    rq_activate_all_grippers(True)
    # end: URCap Program Node
  end
  $ 57 "zero_ftsensor()"
  zero_ftsensor()
  $ 58 "EXTT"
  $ 59 "Set GRP_3F_Enable=Off"
  set_standard_digital_out(4, False)
  $ 60 "Set DO[6]=Off"
  set_standard_digital_out(6, False)
  $ 61 "Set GRP_3F_Decap=Off"
  set_standard_digital_out(3, False)
  $ 62 "Set GRP_3F_Cap=Off"
  set_standard_digital_out(2, False)
  $ 63 "Set GRP_3F_Open=Off"
  set_standard_digital_out(5, False)
  $ 64 "PSE_T≔get_tool_free_pose(dir=[0,0,0.150], move_in_base_frame=True)"
  global PSE_T=get_tool_free_pose(dir=[0,0,0.150], move_in_base_frame=True)
  $ 65 "If is_reachable(Base_const, [PSE_T])"
  if (is_reachable(p[0.0,0.0,0.0,0.0,0.0,0.0], [PSE_T])):
    $ 66 "MoveL"
    $ 67 "PSE_T" "breakAfter"
    movel(PSE_T, a=1.2, v=0.15)
  end
  $ 68 "powder dispensing variable init"
  $ 69 "Start_thread≔ False "
  global Start_thread=  False
  $ 70 "vib_mot_thread≔ False "
  global vib_mot_thread=  False
  $ 71 "kp≔0.0002"
  global kp=0.0002
  $ 72 "ki≔0.001"
  global ki=0.001
  $ 73 "kd≔0.01"
  global kd=0.01
  $ 74 "dt≔0.05"
  global dt=0.05
  $ 75 "Integral_error≔0"
  global Integral_error=0
  $ 76 "current_error≔0"
  global current_error=0
  $ 77 "previous_error≔0"
  global previous_error=0
  $ 78 "tilt_increment≔0"
  global tilt_increment=0
  $ 79 "tilt_angle≔-1"
  global tilt_angle=-1
  $ 80 "diff≔0"
  global diff=0
  $ 81 "current_pose≔get_actual_tcp_pose()"
  global current_pose= get_actual_tcp_pose ()
  $ 896 "Thread_1"
  thread Thread_1():
    while (True):
      $ 897 "If Start_thread≟ True "
      if (Start_thread ==   True  ):
        $ 898 "Weight_value≔get_weight()"
        global Weight_value=get_weight()
        $ 899 "sync()"
        sync()
      end
    end
  end
  threadId_Thread_1 = run Thread_1()
  $ 900 "Thread_2"
  thread Thread_2():
    while (True):
      $ 901 "Loop vib_mot_thread≟ True "
      thread Thread_while_901():
        while (True):
          $ 902 "diff≔Target_weight-Weight_value"
          global diff=Target_weight-Weight_value
          $ 903 "If diff>0.08"
          global thread_flag_903=0
          thread Thread_if_903():
            $ 904 "Set AO[0]=4.0"
            set_standard_analog_out(0, 0.4)
            thread_flag_903 = 1
          end
          if (diff>0.08):
            global thread_handler_903=run Thread_if_903()
            while (thread_flag_903 == 0):
              if not(diff>0.08):
                kill thread_handler_903
                thread_flag_903 = 2
              else:
                sync()
              end
            end
          else:
            thread_flag_903 = 2
          end
          if (thread_flag_903 == 2):
            $ 905 "ElseIf diff≥0.04 and diff≤0.08"
            global thread_flag_905=0
            thread Thread_if_905():
              $ 906 "vibration_1()"
              vibration_1()
              thread_flag_905 = 1
            end
            if (diff >= 0.04 and diff <= 0.08):
              global thread_handler_905=run Thread_if_905()
              while (thread_flag_905 == 0):
                if not(diff >= 0.04 and diff <= 0.08):
                  kill thread_handler_905
                  thread_flag_905 = 2
                else:
                  sync()
                end
              end
            else:
              thread_flag_905 = 2
            end
            if (thread_flag_905 == 2):
              $ 907 "ElseIf diff≥0.01 and diff<0.04"
              if (diff >= 0.01 and diff<0.04):
                $ 908 "vibration_2()"
                vibration_2()
              else:
                $ 909 "ElseIf diff>0 and diff<0.01"
                if (diff>0 and diff<0.01):
                  $ 910 "vibration_3()"
                  vibration_3()
                else:
                  $ 911 "Else" "noBreak"
                  $ 912 "Set AO[0]=0.0"
                  set_standard_analog_out(0, 0.0)
                end
              end
            end
          end
        end
      end
      if (vib_mot_thread ==   True  ):
        global thread_handler_901=run Thread_while_901()
        while (vib_mot_thread ==   True  ):
          sync()
        end
        kill thread_handler_901
      end
      $ 915 "sync()"
      sync()
    end
  end
  threadId_Thread_2 = run Thread_2()
  while (True):
    $ 82 "Robot Program"
    $ 83 "MAIN"
    $ 84 "command_manager(external_control='uGO', cond_suspend=(ITM_Manipulated and AMR_AtTarget and AMR_Charging and AMR_Battery<40), cond_unsuspend=(AMR_Battery≟60))"
    command_manager(external_control="uGO", cond_suspend=(ITM_Manipulated  and  AMR_AtTarget  and  AMR_Charging  and  AMR_Battery<40), cond_unsuspend=(AMR_Battery == 60))
    $ 85 "log_state(STATE_Info)"
    log_state(STATE_Info)
    $ 86 "Switch STATE"
    switch_1 = STATE
    $ 87 "Case 1"
    if (1 == switch_1):
      $ 88 "Stopping"
      $ 89 "STATE_Info≔'Stopping'"
      global STATE_Info="Stopping"
      $ 90 "end_freedrive_mode()"
      end_freedrive_mode()
      $ 91 "Set"
      set_tcp(p[0.0,0.0,0.161,3.1415,0.0,0.0])
      $ 92 "PSE_T≔get_tool_free_pose(dir=[0,0,0.150], move_in_base_frame=True)"
      global PSE_T=get_tool_free_pose(dir=[0,0,0.150], move_in_base_frame=True)
      $ 93 "If is_reachable(Base_const, [PSE_T])"
      if (is_reachable(p[0.0,0.0,0.0,0.0,0.0,0.0], [PSE_T])):
        $ 94 "MoveL"
        $ 95 "PSE_T" "breakAfter"
        movel(PSE_T, a=1.2, v=0.15)
      end
      $ 96 "do_transition(keep_rxry=OBJ_Picked, r=0)"
      do_transition(keep_rxry=OBJ_Picked, r=0)
      $ 105 "Call Sub_AMR_MiR_V3"
      Sub_AMR_MiR_V3()
      $ 106 "If stopping() and AMR_Done"
      if (stopping()  and  AMR_Done):
        $ 107 "STATE≔2"
        global STATE=2
        $ 108 "ugo_update_outputs()"
        ugo_update_outputs()
      end
    elif (2 == switch_1):
      $ 109 "Case 2"
      $ 110 "Stopped"
      $ 111 "STATE_Info≔'Stopped'"
      global STATE_Info="Stopped"
      $ 112 "Call Sub_AMR_MiR_V3"
      Sub_AMR_MiR_V3()
      $ 113 "If CMD_Reset"
      if (CMD_Reset):
        $ 114 "STATE≔3"
        global STATE=3
        $ 115 "ugo_update_outputs()"
        ugo_update_outputs()
      end
    elif (3 == switch_1):
      $ 116 "Case 3"
      $ 117 " Resetting"
      $ 118 "STATE_Info≔'Resetting'"
      global STATE_Info="Resetting"
      $ 119 "uML"
      $ 120 "reset_error()"
      reset_error()
      $ 121 "reset_warning()"
      reset_warning()
      $ 122 "PROCESS_Step≔0"
      global PROCESS_Step=0
      $ 123 "PROCESS_Info≔''"
      global PROCESS_Info=""
      $ 124 "ARM_Referenced≔ False "
      global ARM_Referenced=  False
      $ 125 "WRK_Done≔ False "
      global WRK_Done=  False
      $ 126 "ITM_Prepared≔ False "
      global ITM_Prepared=  False
      $ 127 "ITM_Manipulated≔ False "
      global ITM_Manipulated=  False
      $ 128 "STP≔0"
      global STP=0
      $ 129 "Action≔0"
      global Action=0
      $ 130 "Action_Info≔''"
      global Action_Info=""
      $ 131 "ITM_ID≔0"
      global ITM_ID=0
      $ 132 "JIG≔0"
      global JIG=0
      $ 133 "JIG_Slot≔0"
      global JIG_Slot=0
      $ 134 "Task_info≔''"
      global Task_info=""
      $ 135 "Set"
      set_tcp(p[0.0,0.0,0.161,3.1415,0.0,0.0])
      $ 136 "App"
      $ 137 "'ADD APPLICATION SPECIFIC COMMANDS'"
      # 'ADD APPLICATION SPECIFIC COMMANDS'
      $ 138 "OBJ_Type≔0"
      global OBJ_Type=0
      $ 139 "OBJ_Nbr≔0"
      global OBJ_Nbr=0
      $ 140 "If CNT_Rack_Output≥50"
      if (CNT_Rack_Output >= 50):
        $ 141 "CNT_Rack_Output≔0"
        global CNT_Rack_Output=0
      end
      $ 142 "TASK≔struct(ID=0, NAVI=struct(target=0, footprint=0, protectiveOff=0, dock=0), WORK=struct(ITM_ID_Src=0, JIG_ID_Src=0, OBJ_Nbr_Src=0, ACT_Src=0, ITM_ID_Tgt=0, JIG_ID_Tgt=0, OBJ_Nbr_Tgt=0, ACT_Tgt=0, OBJ_Type=0))"
      global TASK=struct(ID=0, NAVI=struct(target=0, footprint=0, protectiveOff=0, dock=0), WORK=struct(ITM_ID_Src=0, JIG_ID_Src=0, OBJ_Nbr_Src=0, ACT_Src=0, ITM_ID_Tgt=0, JIG_ID_Tgt=0, OBJ_Nbr_Tgt=0, ACT_Tgt=0, OBJ_Type=0))
      $ 143 "Call Sub_AMR_MiR_V3"
      Sub_AMR_MiR_V3()
      $ 144 "If resetting() and AMR_Done"
      if (resetting()  and  AMR_Done):
        $ 145 "STATE≔4"
        global STATE=4
        $ 146 "ugo_update_outputs()"
        ugo_update_outputs()
      end
    elif (4 == switch_1):
      $ 147 "Case 4"
      $ 148 "Idle"
      $ 149 "STATE_Info≔'Idle'"
      global STATE_Info="Idle"
      $ 150 "If CMD_Start"
      if (CMD_Start):
        $ 151 "STATE≔5"
        global STATE=5
        $ 152 "ugo_update_outputs()"
        ugo_update_outputs()
      end
    elif (5 == switch_1):
      $ 153 "Case 5"
      $ 154 "Starting"
      $ 155 "STATE_Info≔'Starting'"
      global STATE_Info="Starting"
      $ 156 "'ADD COMMANDS WHAT TO START WITH'"
      # 'ADD COMMANDS WHAT TO START WITH'
      $ 157 "Call Sub_AMR_MiR_V3"
      Sub_AMR_MiR_V3()
      $ 158 "get ugo data"
      $ 159 "Assign Tasks"
      $ 160 "TASK.ID = ugo_get_task()"
      TASK.ID = ugo_get_task()
      $ 161 "If TASK.ID≟1"
      if (TASK.ID == 1):
        $ 162 "Task_info≔'Charge'"
        global Task_info="Charge"
        $ 163 "Parameters"
        $ 164 "AMR_PosTarget≔1"
        global AMR_PosTarget=1
      else:
        $ 165 "ElseIf TASK.ID≟9"
        if (TASK.ID == 9):
          $ 166 "'Pick Sarstedt Rack from Variable source'"
          # 'Pick Sarstedt Rack from Variable source'
          $ 167 "Task_info≔'Navigate to Target'"
          global Task_info="Navigate to Target"
          $ 168 "Parameters"
          $ 169 "AMR_PosTarget≔UGO.read_input('00','ITM_ID')"
          global AMR_PosTarget=UGO.read_input("00","ITM_ID")
        else:
          $ 170 "ElseIf TASK.ID≟10"
          if (TASK.ID == 10):
            $ 171 "'Pick Sarstedt Rack from Variable source'"
            # 'Pick Sarstedt Rack from Variable source'
            $ 172 "Task_info≔'Pick Rack'"
            global Task_info="Pick Rack"
            $ 173 "AMR_PosTarget≔2"
            global AMR_PosTarget=2
            $ 174 "Parameters"
            $ 175 "ITM_ID≔UGO.read_input('00','ITM_ID')"
            global ITM_ID=UGO.read_input("00","ITM_ID")
            $ 176 "JIG≔UGO.read_input('00','JIG_ID')"
            global JIG=UGO.read_input("00","JIG_ID")
            $ 177 "OBJ_Type≔3"
            global OBJ_Type=3
          else:
            $ 178 "ElseIf TASK.ID≟11"
            if (TASK.ID == 11):
              $ 179 "'Place Sarstedt Rack on Variable target'"
              # 'Place Sarstedt Rack on Variable target'
              $ 180 "Task_info≔'Place Rack'"
              global Task_info="Place Rack"
              $ 181 "AMR_PosTarget≔2"
              global AMR_PosTarget=2
              $ 182 "Parameters"
              $ 183 "ITM_ID≔UGO.read_input('00','ITM_ID')"
              global ITM_ID=UGO.read_input("00","ITM_ID")
              $ 184 "JIG≔UGO.read_input('00','JIG_ID')"
              global JIG=UGO.read_input("00","JIG_ID")
              $ 185 "OBJ_Type≔3"
              global OBJ_Type=3
            else:
              $ 187 "ElseIf TASK.ID≟12"
              if (TASK.ID == 12):
                $ 188 "Task_info≔'Decapping'"
                global Task_info="Decapping"
                $ 189 "Parameters"
                $ 190 "ITM_ID≔1"
                global ITM_ID=1
                $ 191 "AMR_PosTarget≔AMR_PosActual"
                global AMR_PosTarget=AMR_PosActual
                $ 192 "PRC_TubCounter≔0"
                global PRC_TubCounter=0
              else:
                $ 193 "ElseIf TASK.ID≟13"
                if (TASK.ID == 13):
                  $ 194 "Task_info≔'Empty racks'"
                  global Task_info="Empty racks"
                  $ 195 "Parameters"
                  $ 196 "ITM_ID≔1"
                  global ITM_ID=1
                  $ 197 "AMR_PosTarget≔AMR_PosActual"
                  global AMR_PosTarget=AMR_PosActual
                else:
                  $ 198 "ElseIf TASK.ID≟16"
                  if (TASK.ID == 16):
                    $ 199 "Task_info≔'Decap + Barcode'"
                    global Task_info="Decap + Barcode"
                    $ 200 "Parameters"
                    $ 202 "OBJs_String≔UGO.read_input('00','ObjPos')"
                    global OBJs_String=UGO.read_input("00","ObjPos")
                    $ 203 "OBJs_List≔make_list(length = elements_in_string(OBJs_String), initial_value = -1, capacity = 50)"
                    global OBJs_List=make_list(length = elements_in_string(OBJs_String), initial_value = -1, capacity = 50)
                    $ 204 "OBJs_List≔string_to_list(OBJs_String)"
                    global OBJs_List=string_to_list(OBJs_String)
                    $ 205 "ITM_ID≔1"
                    global ITM_ID=1
                    $ 206 "OBJ_Type≔2"
                    global OBJ_Type=2
                    $ 207 "JIG≔7"
                    global JIG=7
                    $ 208 "AMR_PosTarget≔AMR_PosActual"
                    global AMR_PosTarget=AMR_PosActual
                  else:
                    $ 209 "ElseIf TASK.ID≟30"
                    if (TASK.ID == 30):
                      $ 210 "Task_info≔'Getting bottles'"
                      global Task_info="Getting bottles"
                      $ 211 "Parameters"
                      $ 212 "ITM_ID≔1"
                      global ITM_ID=1
                      $ 213 "OBJ_Type≔4"
                      global OBJ_Type=4
                      $ 214 "JIG≔9"
                      global JIG=9
                      $ 215 "AMR_PosTarget≔4"
                      global AMR_PosTarget=4
                    else:
                      $ 216 "ElseIf TASK.ID≟40"
                      if (TASK.ID == 40):
                        $ 217 "Task_info≔'Placing bottles'"
                        global Task_info="Placing bottles"
                        $ 218 "Parameters"
                        $ 219 "ITM_ID≔1"
                        global ITM_ID=1
                        $ 220 "OBJ_Type≔4"
                        global OBJ_Type=4
                        $ 221 "JIG≔10"
                        global JIG=10
                        $ 222 "AMR_PosTarget≔4"
                        global AMR_PosTarget=4
                      else:
                        $ 223 "ElseIf TASK.ID≟41"
                        if (TASK.ID == 41):
                          $ 224 "Task_info≔'Shaking bottle'"
                          global Task_info="Shaking bottle"
                          $ 225 "Parameters"
                          $ 226 "ITM_ID≔1"
                          global ITM_ID=1
                          $ 227 "OBJ_Type≔4"
                          global OBJ_Type=4
                          $ 228 "JIG≔11"
                          global JIG=11
                          $ 229 "AMR_PosTarget≔4"
                          global AMR_PosTarget=4
                        else:
                          $ 230 "ElseIf TASK.ID≟42"
                          if (TASK.ID == 42):
                            $ 231 "Task_info≔'Decap the bottle'"
                            global Task_info="Decap the bottle"
                            $ 232 "Parameters"
                            $ 233 "ITM_ID≔1"
                            global ITM_ID=1
                            $ 234 "OBJ_Type≔4"
                            global OBJ_Type=4
                            $ 235 "AMR_PosTarget≔4"
                            global AMR_PosTarget=4
                          else:
                            $ 236 "ElseIf TASK.ID≟43"
                            if (TASK.ID == 43):
                              $ 237 "Task_info≔'Pick the Rack'"
                              global Task_info="Pick the Rack"
                              $ 238 "AMR_PosTarget≔5"
                              global AMR_PosTarget=5
                              $ 239 "Parameters"
                              $ 240 "ITM_ID≔UGO.read_input('00','ITM_ID')"
                              global ITM_ID=UGO.read_input("00","ITM_ID")
                              $ 241 "JIG≔UGO.read_input('00','JIG_ID')"
                              global JIG=UGO.read_input("00","JIG_ID")
                              $ 242 "OBJ_Type≔3"
                              global OBJ_Type=3
                            else:
                              $ 243 "ElseIf TASK.ID≟45"
                              if (TASK.ID == 45):
                                $ 244 "Task_info≔'pick the Vial'"
                                global Task_info="pick the Vial"
                                $ 245 "Parameters"
                                $ 246 "ITM_ID≔1"
                                global ITM_ID=1
                                $ 247 "OBJ_Type≔4"
                                global OBJ_Type=4
                                $ 248 "JIG≔12"
                                global JIG=12
                                $ 249 "AMR_PosTarget≔5"
                                global AMR_PosTarget=5
                              else:
                                $ 250 "ElseIf TASK.ID≟46"
                                if (TASK.ID == 46):
                                  $ 251 "Task_info≔'Decap the Vial'"
                                  global Task_info="Decap the Vial"
                                  $ 252 "Parameters"
                                  $ 253 "ITM_ID≔1"
                                  global ITM_ID=1
                                  $ 254 "OBJ_Type≔4"
                                  global OBJ_Type=4
                                  $ 255 "JIG≔13"
                                  global JIG=13
                                  $ 256 "AMR_PosTarget≔5"
                                  global AMR_PosTarget=5
                                else:
                                  $ 257 "ElseIf TASK.ID≟47"
                                  if (TASK.ID == 47):
                                    $ 258 "Task_info≔'Liquid Transfer'"
                                    global Task_info="Liquid Transfer"
                                    $ 259 "Parameters"
                                    $ 260 "ITM_ID≔1"
                                    global ITM_ID=1
                                    $ 261 "OBJ_Type≔4"
                                    global OBJ_Type=4
                                    $ 262 "JIG≔14"
                                    global JIG=14
                                    $ 263 "AMR_PosTarget≔3"
                                    global AMR_PosTarget=3
                                  else:
                                    $ 264 "ElseIf TASK.ID≟48"
                                    if (TASK.ID == 48):
                                      $ 265 "Task_info≔'Place_rack'"
                                      global Task_info="Place_rack"
                                      $ 266 "Parameters"
                                      $ 267 "ITM_ID≔1"
                                      global ITM_ID=1
                                      $ 268 "OBJ_Type≔3"
                                      global OBJ_Type=3
                                      $ 269 "JIG≔7"
                                      global JIG=7
                                      $ 270 "AMR_PosTarget≔5"
                                      global AMR_PosTarget=5
                                    else:
                                      $ 271 "ElseIf TASK.ID≟49"
                                      if (TASK.ID == 49):
                                        $ 272 "Task_info≔'Pick Containers'"
                                        global Task_info="Pick Containers"
                                        $ 273 "Parameters"
                                        $ 274 "ITM_ID≔1"
                                        global ITM_ID=1
                                        $ 275 "OBJ_Type≔6"
                                        global OBJ_Type=6
                                        $ 276 "JIG≔15"
                                        global JIG=15
                                        $ 277 "AMR_PosTarget≔3"
                                        global AMR_PosTarget=3
                                      else:
                                        $ 278 "ElseIf TASK.ID≟50"
                                        if (TASK.ID == 50):
                                          $ 279 "Task_info≔'Decap Containers'"
                                          global Task_info="Decap Containers"
                                          $ 280 "Parameters"
                                          $ 281 "ITM_ID≔1"
                                          global ITM_ID=1
                                          $ 282 "OBJ_Type≔6"
                                          global OBJ_Type=6
                                          $ 283 "JIG≔16"
                                          global JIG=16
                                          $ 284 "AMR_PosTarget≔5"
                                          global AMR_PosTarget=5
                                        else:
                                          $ 285 "ElseIf TASK.ID≟51"
                                          if (TASK.ID == 51):
                                            $ 286 "Task_info≔'Detect Spatula and transfer powder'"
                                            global Task_info="Detect Spatula and transfer powder"
                                            $ 287 "Parameters"
                                            $ 288 "ITM_ID≔1"
                                            global ITM_ID=1
                                            $ 289 "Target_weight≔(UGO.read_input('00','Target_weight'))/1000"
                                            global Target_weight=(UGO.read_input("00","Target_weight"))/1000
                                            $ 290 "OBJ_Type≔8"
                                            global OBJ_Type=8
                                            $ 291 "JIG≔16"
                                            global JIG=16
                                            $ 292 "AMR_PosTarget≔5"
                                            global AMR_PosTarget=5
                                          else:
                                            $ 293 "ElseIf TASK.ID≟99"
                                            if (TASK.ID == 99):
                                              $ 294 "Task_info≔'Decapping and barcode alignment'"
                                              global Task_info="Decapping and barcode alignment"
                                              $ 295 "Parameters"
                                              $ 296 "PRC_TubNumber≔UGO.read_input('00','TubesNb')"
                                              global PRC_TubNumber=UGO.read_input("00","TubesNb")
                                              $ 297 "PRC_TubCounter≔0"
                                              global PRC_TubCounter=0
                                              $ 298 "ITM_ID≔1"
                                              global ITM_ID=1
                                              $ 299 "AMR_PosTarget≔AMR_PosActual"
                                              global AMR_PosTarget=AMR_PosActual
                                            else:
                                              $ 334 "Else" "noBreak"
                                              $ 335 "set_error(ERROR_WRONG_ORDER)"
                                              set_error(ERROR_WRONG_ORDER)
                                            end
                                          end
                                        end
                                      end
                                    end
                                  end
                                end
                              end
                            end
                          end
                        end
                      end
                    end
                  end
                end
              end
            end
          end
        end
      end
      $ 336 "test ugo"
      $ 337 "Wait: 0.2"
      sleep(0.2)
      $ 338 "ugo_update_outputs()"
      ugo_update_outputs()
      $ 339 "If starting() and AMR_Done"
      if (starting()  and  AMR_Done):
        $ 340 "log_message(Task_info, 'New Task: ')"
        log_message(Task_info, "New Task: ")
        $ 341 "log_message(to_str(TASK.ID), 'Task_ID: ')"
        log_message(to_str(TASK.ID), "Task_ID: ")
        $ 342 "do_transition(keep_rxry=OBJ_Picked)"
        do_transition(keep_rxry=OBJ_Picked)
        $ 343 "STATE≔6"
        global STATE=6
        $ 344 "ugo_update_outputs()"
        ugo_update_outputs()
      end
    elif (6 == switch_1):
      $ 345 "Case 6"
      $ 346 "Execute"
      $ 347 "STATE_Info≔'Execute'"
      global STATE_Info="Execute"
      $ 348 "If  not CMD_Hold and not CMD_Suspend"
      global thread_flag_348=0
      thread Thread_if_348():
        $ 349 "Switch PROCESS_Step"
        switch_2 = PROCESS_Step
        $ 350 "Case 0"
        if (0 == switch_2):
          $ 351 "PROCESS_Info≔'process control'"
          global PROCESS_Info="process control"
          $ 352 "log_process(PROCESS_Info)"
          log_process(PROCESS_Info)
          $ 353 "process control"
          $ 354 "If  not AMR_AtTarget"
          if (  not  AMR_AtTarget):
            $ 355 "PROCESS_Step≔1"
            global PROCESS_Step=1
          else:
            $ 356 "ElseIf (( not ITM_Prepared and  not WRK_Done) or (ITM_Prepared and WRK_Done))"
            if (((  not  ITM_Prepared  and    not  WRK_Done)  or  (ITM_Prepared  and  WRK_Done))):
              $ 357 "PROCESS_Step≔2"
              global PROCESS_Step=2
            else:
              $ 358 "ElseIf  not WRK_Done"
              if (  not  WRK_Done):
                $ 359 "PROCESS_Step≔3"
                global PROCESS_Step=3
              else:
                $ 360 "Else" "noBreak"
                $ 361 "task finished"
                $ 362 "PROCESS_Info≔''"
                global PROCESS_Info=""
                $ 363 "STATE≔7"
                global STATE=7
                $ 364 "ugo_update_outputs()"
                ugo_update_outputs()
              end
            end
          end
        elif (1 == switch_2):
          $ 365 "Case 1"
          $ 366 "navigate"
          $ 367 "'MOVING THE uML'"
          # 'MOVING THE uML'
          $ 368 "PROCESS_Info≔'move to target'"
          global PROCESS_Info="move to target"
          $ 369 "log_process(PROCESS_Info)"
          log_process(PROCESS_Info)
          $ 370 "If TASK.ID≟1"
          if (TASK.ID == 1):
            $ 371 "Action≔51"
            global Action=51
          else:
            $ 372 "Else" "noBreak"
            $ 373 "Action≔52"
            global Action=52
          end
          $ 374 "Call Sub_AMR_MiR_V3"
          Sub_AMR_MiR_V3()
          $ 375 "If AMR_Done"
          if (AMR_Done):
            $ 376 "PROCESS_Step≔0"
            global PROCESS_Step=0
          end
        elif (2 == switch_2):
          $ 377 "Case 2"
          $ 378 "prepare"
          $ 379 "'THINGS THAT HAVE TO BE DONE ONCE IN A SEQUENCE,WORKFLOW'"
          # 'THINGS THAT HAVE TO BE DONE ONCE IN A SEQUENCE,WORKFLOW'
          $ 380 "PROCESS_Info≔'prepare for work'"
          global PROCESS_Info="prepare for work"
          $ 381 "log_process(PROCESS_Info)"
          log_process(PROCESS_Info)
          $ 382 "If TASK.WORK.ITM_ID_Src>1"
          if (TASK.WORK.ITM_ID_Src>1):
            $ 383 "ITM_ID≔TASK.WORK.ITM_ID_Src"
            global ITM_ID=TASK.WORK.ITM_ID_Src
          else:
            $ 384 "ElseIf TASK.WORK.ITM_ID_Tgt>1"
            if (TASK.WORK.ITM_ID_Tgt>1):
              $ 385 "ITM_ID≔TASK.WORK.ITM_ID_Tgt"
              global ITM_ID=TASK.WORK.ITM_ID_Tgt
            end
          end
          $ 386 "If  not ARM_Referenced and (ITM_ID≠0)"
          if (  not  ARM_Referenced  and  (ITM_ID != 0)):
            $ 387 "STP≔1"
            global STP=1
          else:
            $ 388 "ElseIf ARM_Referenced or (ITM_ID≟0)"
            if (ARM_Referenced  or  (ITM_ID == 0)):
              $ 389 "STP≔2"
              global STP=2
            end
          end
          $ 390 "Switch STP"
          switch_3 = STP
          $ 391 "Case 1"
          if (1 == switch_3):
            $ 392 "reference"
            $ 393 "STP_Info≔'reference at target position'"
            global STP_Info="reference at target position"
            $ 394 "log_step(STP_Info)"
            log_step(STP_Info)
            $ 395 "If ITM_ID≟1"
            if (ITM_ID == 1):
              $ 396 "CAM_Done≔ True "
              global CAM_Done=  True
            else:
              $ 397 "Else" "noBreak"
              $ 398 "Action≔131"
              global Action=131
              $ 399 "Call Sub_Vision_V18"
              Sub_Vision_V18()
            end
            $ 401 "If CAM_Done and  not ERROR.FLAG"
            if (CAM_Done  and    not  ERROR.FLAG):
              $ 402 "log_step('ARM referenced')"
              log_step("ARM referenced")
              $ 403 "ARM_Referenced≔ True "
              global ARM_Referenced=  True
            end
          elif (2 == switch_3):
            $ 404 "Case 2"
            $ 405 "manipulate"
            $ 406 "STP_Info≔'manipulate item'"
            global STP_Info="manipulate item"
            $ 407 "log_step(STP_Info)"
            log_step(STP_Info)
            $ 408 "'In case pressing button is needed'"
            # 'In case pressing button is needed'
            $ 409 "If found_in_list(ITM_ID, ITM_ID_List)"
            if (found_in_list(ITM_ID, ITM_ID_List)):
              $ 410 "Switch ITM_ID"
              switch_4 = ITM_ID
              $ 411 "Case 0"
              if (0 == switch_4):
                $ 412 "ITM_Manipulated≔ not ITM_Manipulated"
                global ITM_Manipulated=  not  ITM_Manipulated
              elif (1 == switch_4):
                $ 413 "Case 1"
                $ 414 "ITM_Manipulated≔ not ITM_Manipulated"
                global ITM_Manipulated=  not  ITM_Manipulated
              elif (2 == switch_4):
                $ 415 "Case 2"
              else:
                $ 425 "Default Case"
                $ 426 "ITM_Manipulated≔ not ITM_Manipulated"
                global ITM_Manipulated=  not  ITM_Manipulated
              end
            end
          end
          $ 427 "ITM_Prepared≔(ITM_Manipulated or  not found_in_list(ITM_ID, ITM_ID_List)) and (ARM_Referenced or ITM_ID≟0) and  not WRK_Done"
          global ITM_Prepared=(ITM_Manipulated  or    not  found_in_list(ITM_ID, ITM_ID_List))  and  (ARM_Referenced  or  ITM_ID == 0)  and    not  WRK_Done
          $ 428 "STP≔0"
          global STP=0
          $ 429 "STP_Info≔''"
          global STP_Info=""
          $ 430 "PROCESS_Step≔0"
          global PROCESS_Step=0
        elif (3 == switch_2):
          $ 431 "Case 3"
          $ 432 "work"
          $ 433 "'ADD EVERY MACHINE, OBJECT, STATION TO WORK ON'"
          # 'ADD EVERY MACHINE, OBJECT, STATION TO WORK ON'
          $ 434 "Switch ITM_ID"
          switch_3 = ITM_ID
          $ 435 "Case 1"
          if (1 == switch_3):
            $ 436 "uLM"
            $ 437 "If TASK.ID≟12"
            if (TASK.ID == 12):
              $ 438 "fill racks"
              $ 439 "Action≔151"
              global Action=151
              $ 440 "Call Sub_Vision_V18"
              Sub_Vision_V18()
              $ 441 "If  not ERROR.FLAG"
              if (  not  ERROR.FLAG):
                $ 442 "Actions for the task"
                $ 443 "Action≔1"
                global Action=1
                $ 444 "JIG≔2"
                global JIG=2
                $ 445 "JIG_Slot≔CAM_Result[0]"
                global JIG_Slot=CAM_Result[0]
                $ 446 "OBJ_Nbr≔CAM_Result[0]"
                global OBJ_Nbr=CAM_Result[0]
                $ 447 "OBJ_Type≔2"
                global OBJ_Type=2
                $ 448 "Call Sub_Action_V4"
                Sub_Action_V4()
                $ 449 "If OBJ_Picked"
                if (OBJ_Picked):
                  $ 450 "CAM_Result.remove(0)"
                  CAM_Result.remove(0)
                  $ 451 "PRC_TubCounter≔PRC_TubCounter+1"
                  global PRC_TubCounter=PRC_TubCounter+1
                  $ 452 "If PRC_TubCounter%4≟0"
                  if (PRC_TubCounter%4 == 0):
                    $ 453 "JIG_Slot≔4"
                    global JIG_Slot=4
                  else:
                    $ 454 "Else" "noBreak"
                    $ 455 "JIG_Slot≔PRC_TubCounter%4"
                    global JIG_Slot=PRC_TubCounter%4
                  end
                  $ 456 "OBJ_Nbr≔ceil(PRC_TubCounter/4)"
                  global OBJ_Nbr=ceil(PRC_TubCounter/4)
                  $ 457 "Action≔2"
                  global Action=2
                  $ 458 "JIG≔4"
                  global JIG=4
                  $ 459 "Call Sub_Action_V4"
                  Sub_Action_V4()
                  $ 460 "Action≔151"
                  global Action=151
                  $ 461 "Call Sub_Vision_V18"
                  Sub_Vision_V18()
                end
              end
              $ 462 "If (CAM_Captures≥CAM_PRM_Retries) or (PRC_TubCounter≥32)"
              if ((CAM_Captures >= CAM_PRM_Retries)  or  (PRC_TubCounter >= 32)):
                $ 463 "PROCESS_Step≔0"
                global PROCESS_Step=0
                $ 464 "WRK_Done≔ True "
                global WRK_Done=  True
              end
            else:
              $ 465 "ElseIf TASK.ID≟10"
              if (TASK.ID == 10):
                $ 466 "Pick Rack"
                $ 467 "Action≔131"
                global Action=131
                $ 468 "Call Sub_Vision_V18"
                Sub_Vision_V18()
                $ 469 "Action≔1"
                global Action=1
                $ 470 "Call Sub_Action_V4"
                Sub_Action_V4()
                $ 471 "PROCESS_Step≔0"
                global PROCESS_Step=0
                $ 472 "WRK_Done≔ True "
                global WRK_Done=  True
              else:
                $ 473 "ElseIf TASK.ID≟11"
                if (TASK.ID == 11):
                  $ 474 "Place Rack"
                  $ 475 "Action≔2"
                  global Action=2
                  $ 476 "Call Sub_Action_V4"
                  Sub_Action_V4()
                  $ 477 "PROCESS_Step≔0"
                  global PROCESS_Step=0
                  $ 478 "WRK_Done≔ True "
                  global WRK_Done=  True
                else:
                  $ 479 "ElseIf TASK.ID≟13"
                  if (TASK.ID == 13):
                    $ 480 "empty racks"
                    $ 481 "pick"
                    $ 482 "Action≔1"
                    global Action=1
                    $ 483 "JIG≔4"
                    global JIG=4
                    $ 484 "If PRC_TubCounter%4≟0"
                    if (PRC_TubCounter%4 == 0):
                      $ 485 "JIG_Slot≔4"
                      global JIG_Slot=4
                    else:
                      $ 486 "Else" "noBreak"
                      $ 487 "JIG_Slot≔PRC_TubCounter%4"
                      global JIG_Slot=PRC_TubCounter%4
                    end
                    $ 488 "OBJ_Nbr≔ceil(PRC_TubCounter/4)"
                    global OBJ_Nbr=ceil(PRC_TubCounter/4)
                    $ 489 "OBJ_Type≔2"
                    global OBJ_Type=2
                    $ 490 "Call Sub_Action_V4"
                    Sub_Action_V4()
                    $ 491 "If OBJ_Picked"
                    if (OBJ_Picked):
                      $ 492 "Action≔2"
                      global Action=2
                      $ 493 "JIG≔3"
                      global JIG=3
                      $ 494 "JIG_Slot≔1"
                      global JIG_Slot=1
                      $ 495 "CNT_Rack_Output≔CNT_Rack_Output + 1"
                      global CNT_Rack_Output=CNT_Rack_Output + 1
                      $ 496 "OBJ_Nbr≔CNT_Rack_Output"
                      global OBJ_Nbr=CNT_Rack_Output
                      $ 497 "Call Sub_Action_V4"
                      Sub_Action_V4()
                      $ 498 "If  not ERROR.FLAG"
                      if (  not  ERROR.FLAG):
                        $ 499 "PRC_TubCounter≔PRC_TubCounter - 1"
                        global PRC_TubCounter=PRC_TubCounter - 1
                      end
                    end
                    $ 500 "If CNT_Rack_Output≥50 or PRC_TubCounter≤0"
                    if (CNT_Rack_Output >= 50  or  PRC_TubCounter <= 0):
                      $ 501 "PROCESS_Step≔0"
                      global PROCESS_Step=0
                      $ 502 "WRK_Done≔ True "
                      global WRK_Done=  True
                    end
                  else:
                    $ 503 "ElseIf TASK.ID≟16"
                    if (TASK.ID == 16):
                      $ 504 "CAM_Result≔OBJs_List"
                      global CAM_Result=OBJs_List
                      $ 505 "PRC_CntDetect≔0"
                      global PRC_CntDetect=0
                      $ 506 "Loop PRC_CntDetect<CAM_Result.length()"
                      while (PRC_CntDetect<CAM_Result.length()):
                        $ 507 "Action≔1"
                        global Action=1
                        $ 508 "ITM_ID≔1"
                        global ITM_ID=1
                        $ 509 "JIG≔2"
                        global JIG=2
                        $ 510 "OBJ_Type≔2"
                        global OBJ_Type=2
                        $ 511 "JIG_Slot≔CAM_Result[PRC_CntDetect]"
                        global JIG_Slot=CAM_Result[PRC_CntDetect]
                        $ 512 "OBJ_Nbr≔CAM_Result[PRC_CntDetect]"
                        global OBJ_Nbr=CAM_Result[PRC_CntDetect]
                        $ 513 "Call Sub_Action_V4"
                        Sub_Action_V4()
                        $ 514 "JIG≔1"
                        global JIG=1
                        $ 515 "Action≔11"
                        global Action=11
                        $ 516 "Call Sub_Action_V4"
                        Sub_Action_V4()
                        $ 517 "Action≔12"
                        global Action=12
                        $ 518 "Call Sub_Action_V4"
                        Sub_Action_V4()
                        $ 519 "Action≔6"
                        global Action=6
                        $ 520 "JIG≔6"
                        global JIG=6
                        $ 521 "Call Sub_Action_V4"
                        Sub_Action_V4()
                        $ 522 "Action≔13"
                        global Action=13
                        $ 523 "Call Sub_Action_V4"
                        Sub_Action_V4()
                        $ 524 "Action≔1"
                        global Action=1
                        $ 525 "JIG≔1"
                        global JIG=1
                        $ 526 "Call Sub_Action_V4"
                        Sub_Action_V4()
                        $ 527 "If OBJ_Brc_OK"
                        if (OBJ_Brc_OK):
                          $ 528 "JIG≔2"
                          global JIG=2
                          $ 529 "Action≔2"
                          global Action=2
                          $ 530 "OBJ_Nbr≔CAM_Result[PRC_CntDetect]"
                          global OBJ_Nbr=CAM_Result[PRC_CntDetect]
                          $ 531 "JIG_Slot≔CAM_Result[PRC_CntDetect]"
                          global JIG_Slot=CAM_Result[PRC_CntDetect]
                          $ 532 "OBJ_Type≔2"
                          global OBJ_Type=2
                          $ 533 "Call Sub_Action_V4"
                          Sub_Action_V4()
                        else:
                          $ 534 "Else" "noBreak"
                          $ 535 "Action≔2"
                          global Action=2
                          $ 536 "JIG≔8"
                          global JIG=8
                          $ 537 "Call Sub_Action_V4"
                          Sub_Action_V4()
                        end
                        $ 538 "PRC_CntDetect≔PRC_CntDetect+1"
                        global PRC_CntDetect=PRC_CntDetect+1
                      end
                      $ 539 "PROCESS_Step≔0"
                      global PROCESS_Step=0
                      $ 540 "WRK_Done≔ True "
                      global WRK_Done=  True
                    else:
                      $ 541 "ElseIf TASK.ID≟30"
                      if (TASK.ID == 30):
                        $ 542 "Pick Bottle"
                        $ 543 "Action≔1"
                        global Action=1
                        $ 544 "Call Sub_Action_V4"
                        Sub_Action_V4()
                        $ 545 "PROCESS_Step≔0"
                        global PROCESS_Step=0
                        $ 546 "WRK_Done≔ True "
                        global WRK_Done=  True
                      else:
                        $ 547 "ElseIf TASK.ID≟40"
                        if (TASK.ID == 40):
                          $ 548 "Place Bottle"
                          $ 549 "Action≔2"
                          global Action=2
                          $ 550 "Call Sub_Action_V4"
                          Sub_Action_V4()
                          $ 551 "PROCESS_Step≔0"
                          global PROCESS_Step=0
                          $ 552 "WRK_Done≔ True "
                          global WRK_Done=  True
                        else:
                          $ 553 "ElseIf TASK.ID≟45"
                          if (TASK.ID == 45):
                            $ 554 "Pick Vial"
                            $ 555 "Action≔31"
                            global Action=31
                            $ 556 "Call Sub_Action_V4"
                            Sub_Action_V4()
                            $ 557 "PROCESS_Step≔0"
                            global PROCESS_Step=0
                            $ 558 "WRK_Done≔ True "
                            global WRK_Done=  True
                          else:
                            $ 559 "ElseIf TASK.ID≟46"
                            if (TASK.ID == 46):
                              $ 560 "Decap Vial"
                              $ 561 "Action≔32"
                              global Action=32
                              $ 562 "Call Sub_Action_V4"
                              Sub_Action_V4()
                              $ 563 "PROCESS_Step≔0"
                              global PROCESS_Step=0
                              $ 564 "WRK_Done≔ True "
                              global WRK_Done=  True
                            else:
                              $ 565 "ElseIf TASK.ID≟47"
                              if (TASK.ID == 47):
                                $ 566 "Liquid transfer"
                                $ 567 "Action≔33"
                                global Action=33
                                $ 568 "Call Sub_Action_V4"
                                Sub_Action_V4()
                                $ 569 "PROCESS_Step≔0"
                                global PROCESS_Step=0
                                $ 570 "WRK_Done≔ True "
                                global WRK_Done=  True
                              else:
                                $ 571 "ElseIf TASK.ID≟48"
                                if (TASK.ID == 48):
                                  $ 572 "Place Rack"
                                  $ 573 "Action≔34"
                                  global Action=34
                                  $ 574 "Call Sub_Action_V4"
                                  Sub_Action_V4()
                                  $ 575 "PROCESS_Step≔0"
                                  global PROCESS_Step=0
                                  $ 576 "WRK_Done≔ True "
                                  global WRK_Done=  True
                                else:
                                  $ 577 "ElseIf TASK.ID≟49"
                                  if (TASK.ID == 49):
                                    $ 578 "Pick Powder container"
                                    $ 579 "Action≔131"
                                    global Action=131
                                    $ 580 "Call Sub_Vision_V18"
                                    Sub_Vision_V18()
                                    $ 583 "Action≔35"
                                    global Action=35
                                    $ 584 "Call Sub_Action_V4"
                                    Sub_Action_V4()
                                    $ 585 "PROCESS_Step≔0"
                                    global PROCESS_Step=0
                                    $ 586 "WRK_Done≔ True "
                                    global WRK_Done=  True
                                  else:
                                    $ 587 "ElseIf TASK.ID≟41"
                                    if (TASK.ID == 41):
                                      $ 588 "shake Bottle"
                                      $ 589 "Action≔30"
                                      global Action=30
                                      $ 590 "Call Sub_Action_V4"
                                      Sub_Action_V4()
                                      $ 591 "PROCESS_Step≔0"
                                      global PROCESS_Step=0
                                      $ 592 "WRK_Done≔ True "
                                      global WRK_Done=  True
                                    else:
                                      $ 593 "ElseIf TASK.ID≟42"
                                      if (TASK.ID == 42):
                                        $ 594 "decap the bottle"
                                        $ 595 "Action≔1"
                                        global Action=1
                                        $ 596 "JIG≔9"
                                        global JIG=9
                                        $ 597 "Call Sub_Action_V4"
                                        Sub_Action_V4()
                                        $ 598 "Action≔11"
                                        global Action=11
                                        $ 599 "JIG≔1"
                                        global JIG=1
                                        $ 600 "Call Sub_Action_V4"
                                        Sub_Action_V4()
                                        $ 601 "Action≔12"
                                        global Action=12
                                        $ 602 "JIG≔1"
                                        global JIG=1
                                        $ 603 "Call Sub_Action_V4"
                                        Sub_Action_V4()
                                        $ 604 "Action≔2"
                                        global Action=2
                                        $ 605 "JIG≔8"
                                        global JIG=8
                                        $ 606 "Call Sub_Action_V4"
                                        Sub_Action_V4()
                                        $ 607 "PROCESS_Step≔0"
                                        global PROCESS_Step=0
                                        $ 608 "WRK_Done≔ True "
                                        global WRK_Done=  True
                                      else:
                                        $ 609 "ElseIf TASK.ID≟43"
                                        if (TASK.ID == 43):
                                          $ 610 "Pick the rack"
                                          $ 611 "Action≔131"
                                          global Action=131
                                          $ 612 "Call Sub_Vision_V18"
                                          Sub_Vision_V18()
                                          $ 613 "Action≔1"
                                          global Action=1
                                          $ 614 "Call Sub_Action_V4"
                                          Sub_Action_V4()
                                          $ 615 "PROCESS_Step≔0"
                                          global PROCESS_Step=0
                                          $ 616 "WRK_Done≔ True "
                                          global WRK_Done=  True
                                        else:
                                          $ 617 "ElseIf TASK.ID≟50"
                                          if (TASK.ID == 50):
                                            $ 618 "Decap containers"
                                            $ 619 "Action≔36"
                                            global Action=36
                                            $ 620 "Call Sub_Action_V4"
                                            Sub_Action_V4()
                                            $ 621 "PROCESS_Step≔0"
                                            global PROCESS_Step=0
                                            $ 622 "WRK_Done≔ True "
                                            global WRK_Done=  True
                                          else:
                                            $ 623 "ElseIf TASK.ID≟51"
                                            if (TASK.ID == 51):
                                              $ 624 "Detect Spatula and transfer powder"
                                              $ 625 "Action≔131"
                                              global Action=131
                                              $ 626 "Call Sub_Vision_V18"
                                              Sub_Vision_V18()
                                              $ 627 "Action≔37"
                                              global Action=37
                                              $ 628 "Call Sub_Action_V4"
                                              Sub_Action_V4()
                                              $ 629 "PROCESS_Step≔0"
                                              global PROCESS_Step=0
                                              $ 630 "WRK_Done≔ True "
                                              global WRK_Done=  True
                                            end
                                          end
                                        end
                                      end
                                    end
                                  end
                                end
                              end
                            end
                          end
                        end
                      end
                    end
                  end
                end
              end
            end
          elif (2 == switch_3):
            $ 631 "Case 2"
          elif (5 == switch_3):
            $ 673 "Case 5"
            $ 674 "SarstedtTable"
            $ 675 "Action≔131"
            global Action=131
            $ 676 "Call Sub_Vision_V18"
            Sub_Vision_V18()
            $ 677 "Action≔1"
            global Action=1
            $ 678 "Call Sub_Action_V4"
            Sub_Action_V4()
            $ 679 "PROCESS_Step≔0"
            global PROCESS_Step=0
            $ 680 "WRK_Done≔ True "
            global WRK_Done=  True
          elif (20 == switch_3):
            $ 681 "Case 20"
          elif (43 == switch_3):
            $ 743 "Case 43"
            $ 744 "Pick the rack"
            $ 745 "Action≔131"
            global Action=131
            $ 746 "Call Sub_Vision_V18"
            Sub_Vision_V18()
            $ 747 "Action≔1"
            global Action=1
            $ 748 "Call Sub_Action_V4"
            Sub_Action_V4()
            $ 749 "PROCESS_Step≔0"
            global PROCESS_Step=0
            $ 750 "WRK_Done≔ True "
            global WRK_Done=  True
          else:
            $ 751 "Default Case"
            $ 752 "WRK_Done≔ True "
            global WRK_Done=  True
            $ 753 "PROCESS_Step≔0"
            global PROCESS_Step=0
          end
        end
        thread_flag_348 = 1
      end
      if (  not  CMD_Hold and not CMD_Suspend):
        global thread_handler_348=run Thread_if_348()
        while (thread_flag_348 == 0):
          if not(  not  CMD_Hold and not CMD_Suspend):
            kill thread_handler_348
            thread_flag_348 = 2
          else:
            sync()
          end
        end
      else:
        thread_flag_348 = 2
      end
      $ 754 "If CMD_Hold"
      if (CMD_Hold):
        $ 755 "STATE≔9"
        global STATE=9
        $ 756 "ugo_update_outputs()"
        ugo_update_outputs()
      else:
        $ 757 "ElseIf CMD_Suspend"
        if (CMD_Suspend):
          $ 758 "STATE≔12"
          global STATE=12
          $ 759 "ugo_update_outputs()"
          ugo_update_outputs()
        end
      end
    elif (7 == switch_1):
      $ 760 "Case 7"
      $ 761 "Completing"
      $ 762 "STATE_Info≔'Completing'"
      global STATE_Info="Completing"
      $ 763 "'ADD COMMANDS FOR COMPLETING THE PROCESS'"
      # 'ADD COMMANDS FOR COMPLETING THE PROCESS'
      $ 764 "do_transition(keep_rxry=OBJ_Picked)"
      do_transition(keep_rxry=OBJ_Picked)
      $ 765 "Call Sub_AMR_MiR_V3"
      Sub_AMR_MiR_V3()
      $ 766 "If completing() and AMR_Done"
      if (completing()  and  AMR_Done):
        $ 767 "STATE≔8"
        global STATE=8
        $ 768 "ugo_update_outputs()"
        ugo_update_outputs()
      end
    elif (8 == switch_1):
      $ 769 "Case 8"
      $ 770 "Complete"
      $ 771 "STATE_Info≔'Complete'"
      global STATE_Info="Complete"
      $ 772 "If CMD_Reset"
      if (CMD_Reset):
        $ 773 "STATE≔3"
        global STATE=3
        $ 774 "ugo_update_outputs()"
        ugo_update_outputs()
      end
    elif (9 == switch_1):
      $ 775 "Case 9"
      $ 776 "Holding"
      $ 777 "STATE_Info≔'Holding'"
      global STATE_Info="Holding"
      $ 778 "stopl(0.5)"
      stopl(0.5)
      $ 779 "Call Sub_AMR_MiR_V3"
      Sub_AMR_MiR_V3()
      $ 780 "If holding() and AMR_Done"
      if (holding()  and  AMR_Done):
        $ 781 "STATE≔10"
        global STATE=10
        $ 782 "ugo_update_outputs()"
        ugo_update_outputs()
      end
    elif (10 == switch_1):
      $ 783 "Case 10"
      $ 784 "Held"
      $ 785 "STATE_Info≔'Held'"
      global STATE_Info="Held"
      $ 786 "If CMD_Unhold"
      if (CMD_Unhold):
        $ 787 "end_freedrive_mode()"
        end_freedrive_mode()
        $ 788 "STATE≔11"
        global STATE=11
        $ 789 "ugo_update_outputs()"
        ugo_update_outputs()
      else:
        $ 790 "ElseIf FNC_Freedrive"
        if (FNC_Freedrive):
          $ 791 "freedrive_mode()"
          freedrive_mode()
        else:
          $ 792 "Else" "noBreak"
          $ 793 "end_freedrive_mode()"
          end_freedrive_mode()
        end
      end
    elif (11 == switch_1):
      $ 794 "Case 11"
      $ 795 "Unholding"
      $ 796 "STATE_Info≔'Unholding'"
      global STATE_Info="Unholding"
      $ 797 "Clearing"
      $ 798 "Switch ERROR.ID"
      switch_2 = ERROR.ID
      $ 799 "Case 1002"
      if (1002 == switch_2):
        $ 800 "AMR_AtTarget≔ False "
        global AMR_AtTarget=  False
        $ 801 "ARM_Referenced≔ False "
        global ARM_Referenced=  False
        $ 802 "ITM_Prepared≔ False "
        global ITM_Prepared=  False
        $ 803 "PROCESS_Step≔1"
        global PROCESS_Step=1
      elif (2007 == switch_2):
        $ 804 "Case 2007"
        $ 805 "PROCESS_Step≔1"
        global PROCESS_Step=1
      end
      $ 806 "reset_error()"
      reset_error()
      $ 807 "reset_warning()"
      reset_warning()
      $ 808 "OBJ_Picked≔gripper_has_object()"
      global OBJ_Picked=gripper_has_object()
      $ 809 "Call Sub_AMR_MiR_V3"
      Sub_AMR_MiR_V3()
      $ 810 "If unholding() and AMR_Done"
      if (unholding()  and  AMR_Done):
        $ 811 "STATE≔6"
        global STATE=6
        $ 812 "ugo_update_outputs()"
        ugo_update_outputs()
      end
    elif (12 == switch_1):
      $ 813 "Case 12"
      $ 814 "Suspending"
      $ 815 "STATE_Info≔'Suspending'"
      global STATE_Info="Suspending"
      $ 816 "PROCESS_Info≔str_cat(PROCESS_Info, ' suspended')"
      global PROCESS_Info=str_cat(PROCESS_Info, " suspended")
      $ 817 "If suspending()"
      if (suspending()):
        $ 818 "STATE≔13"
        global STATE=13
        $ 819 "ugo_update_outputs()"
        ugo_update_outputs()
      end
    elif (13 == switch_1):
      $ 820 "Case 13"
      $ 821 "Suspended"
      $ 822 "STATE_Info≔'Suspended'"
      global STATE_Info="Suspended"
      $ 823 "Call Sub_AMR_MiR_V3"
      Sub_AMR_MiR_V3()
      $ 824 "If CMD_Unsuspend"
      if (CMD_Unsuspend):
        $ 825 "STATE≔14"
        global STATE=14
        $ 826 "ugo_update_outputs()"
        ugo_update_outputs()
      end
    elif (14 == switch_1):
      $ 827 "Case 14"
      $ 828 "Unsuspending"
      $ 829 "STATE_Info≔'Unsuspending'"
      global STATE_Info="Unsuspending"
      $ 830 "PROCESS_Step≔0"
      global PROCESS_Step=0
      $ 831 "If unsuspending()"
      if (unsuspending()):
        $ 832 "STATE≔6"
        global STATE=6
        $ 833 "ugo_update_outputs()"
        ugo_update_outputs()
      end
    elif (15 == switch_1):
      $ 834 "Case 15"
      $ 835 "Aborting"
      $ 836 "STATE_Info≔'Aborting'"
      global STATE_Info="Aborting"
      $ 837 "If aborting()"
      if (aborting()):
        $ 838 "STATE≔16"
        global STATE=16
        $ 839 "ugo_update_outputs()"
        ugo_update_outputs()
      end
    elif (16 == switch_1):
      $ 840 "Case 16"
      $ 841 "Aborted"
      $ 842 "STATE_Info≔'Aborted'"
      global STATE_Info="Aborted"
      $ 843 "If CMD_Clear"
      if (CMD_Clear):
        $ 844 "STATE≔17"
        global STATE=17
        $ 845 "ugo_update_outputs()"
        ugo_update_outputs()
      end
    elif (17 == switch_1):
      $ 846 "Case 17"
      $ 847 "Clearing"
      $ 848 "STATE_Info≔'Clearing'"
      global STATE_Info="Clearing"
      $ 849 "Clearing"
      $ 850 "reset_warning()"
      reset_warning()
      $ 851 "reset_error()"
      reset_error()
      $ 852 "If clearing()"
      if (clearing()):
        $ 853 "STATE≔2"
        global STATE=2
        $ 854 "ugo_update_outputs()"
        ugo_update_outputs()
      end
    end
    $ 855 "log_state(STATE_Info)"
    log_state(STATE_Info)
    $ 856 "log_warning(WARNING.MSG)"
    log_warning(WARNING.MSG)
    $ 857 "log_error(ERROR.MSG)"
    log_error(ERROR.MSG)
    $ 858 "Times"
    $ 859 "Switch STATE"
    switch_1 = STATE
    $ 860 "Case 1"
    if (1 == switch_1):
      $ 861 "TM_St_Stopping≔get_time(STATE_Times[STATE-1])"
      global TM_St_Stopping=get_time(STATE_Times[STATE-1])
    elif (2 == switch_1):
      $ 862 "Case 2"
      $ 863 "TM_St_Stopped≔get_time(STATE_Times[STATE-1])"
      global TM_St_Stopped=get_time(STATE_Times[STATE-1])
    elif (3 == switch_1):
      $ 864 "Case 3"
      $ 865 "TM_St_Resetting≔get_time(STATE_Times[STATE-1])"
      global TM_St_Resetting=get_time(STATE_Times[STATE-1])
    elif (4 == switch_1):
      $ 866 "Case 4"
      $ 867 "TM_St_Idle≔get_time(STATE_Times[STATE-1])"
      global TM_St_Idle=get_time(STATE_Times[STATE-1])
    elif (5 == switch_1):
      $ 868 "Case 5"
      $ 869 "TM_St_Starting≔get_time(STATE_Times[STATE-1])"
      global TM_St_Starting=get_time(STATE_Times[STATE-1])
    elif (6 == switch_1):
      $ 870 "Case 6"
      $ 871 "TM_St_Execute≔get_time(STATE_Times[STATE-1])"
      global TM_St_Execute=get_time(STATE_Times[STATE-1])
    elif (7 == switch_1):
      $ 872 "Case 7"
      $ 873 "TM_St_Completin≔get_time(STATE_Times[STATE-1])"
      global TM_St_Completin=get_time(STATE_Times[STATE-1])
    elif (8 == switch_1):
      $ 874 "Case 8"
      $ 875 "TM_St_Complete≔get_time(STATE_Times[STATE-1])"
      global TM_St_Complete=get_time(STATE_Times[STATE-1])
    elif (9 == switch_1):
      $ 876 "Case 9"
      $ 877 "TM_St_Holding≔get_time(STATE_Times[STATE-1])"
      global TM_St_Holding=get_time(STATE_Times[STATE-1])
    elif (10 == switch_1):
      $ 878 "Case 10"
      $ 879 "TM_St_Held≔get_time(STATE_Times[STATE-1])"
      global TM_St_Held=get_time(STATE_Times[STATE-1])
    elif (11 == switch_1):
      $ 880 "Case 11"
      $ 881 "TM_St_Unholding≔get_time(STATE_Times[STATE-1])"
      global TM_St_Unholding=get_time(STATE_Times[STATE-1])
    elif (12 == switch_1):
      $ 882 "Case 12"
      $ 883 "TM_St_Suspendin≔get_time(STATE_Times[STATE-1])"
      global TM_St_Suspendin=get_time(STATE_Times[STATE-1])
    elif (13 == switch_1):
      $ 884 "Case 13"
      $ 885 "TM_St_Suspended≔get_time(STATE_Times[STATE-1])"
      global TM_St_Suspended=get_time(STATE_Times[STATE-1])
    elif (14 == switch_1):
      $ 886 "Case 14"
      $ 887 "TM_St_Unsuspend≔get_time(STATE_Times[STATE-1])"
      global TM_St_Unsuspend=get_time(STATE_Times[STATE-1])
    elif (15 == switch_1):
      $ 888 "Case 15"
      $ 889 "TM_St_Aborting≔get_time(STATE_Times[STATE-1])"
      global TM_St_Aborting=get_time(STATE_Times[STATE-1])
    elif (16 == switch_1):
      $ 890 "Case 16"
      $ 891 "TM_St_Aborted≔get_time(STATE_Times[STATE-1])"
      global TM_St_Aborted=get_time(STATE_Times[STATE-1])
    elif (17 == switch_1):
      $ 892 "Case 17"
      $ 893 "TM_St_Clearing≔get_time(STATE_Times[STATE-1])"
      global TM_St_Clearing=get_time(STATE_Times[STATE-1])
    end
    $ 895 "Wait: 0.1"
    sleep(0.1)
  end
end
